(* IEC 61131-3 sources: tsplc/packages/vscode-extension/tests/fixtures/conveyor/transport/FB_Conveyor, 1 file *)

(* ---- FB_Conveyor.declaration.st ---- *)
FUNCTION_BLOCK FB_Conveyor
VAR_IN_OUT
	Conveyor : ST_Conveyor;
END_VAR
VAR
	pConveyor : POINTER TO ST_Conveyor;
END_VAR
